(* PLC project g_two_hand_fb_type_i, Anonymous Benchmark Suite 1.0 *)
(* stored: creationDateTime 2026-08-28T00:00:00 *)

FUNCTION_BLOCK TwoHandII
  VAR_INPUT
    LH : BOOL;
    RH : BOOL;
  END_VAR
  VAR_OUTPUT
    Stroke : BOOL;
  END_VAR
  VAR
    BothOff : BOOL;
    Armed : BOOL;
  END_VAR

Stroke := LH AND RH;
END_FUNCTION_BLOCK

PROGRAM g_two_hand_fb_type_i
  VAR_INPUT
    LH : BOOL;
    RH : BOOL;
  END_VAR
  VAR_OUTPUT
    Stroke : BOOL;
  END_VAR
  VAR
    THC0 : TwoHandII;
  END_VAR

(* LD diagram, written out as Structured Text *)
THC0(LH := LH, RH := RH);
Stroke := THC0.Stroke;
END_PROGRAM

CONFIGURATION Config0
  RESOURCE Res0 ON PLC
    TASK tcyclic(INTERVAL := T#10ms, PRIORITY := 0);
    PROGRAM inst0 WITH tcyclic : g_two_hand_fb_type_i;
  END_RESOURCE
END_CONFIGURATION
